FUNCTION_BLOCK AI_LAST_2 (* MERGE 2 AI in 1 AI (LAST WRITER WINS, generic FB) - welcher Socket zuletzt geschrieben hat, gewinnt und wird sofort an OUT durchgereicht *)
  (* Standard: 61499-2; Description: Copyright (c) 2026 Meisterschulen am Ostbahnhof This program and the accompanying materials are made available under the terms of the Eclipse Public License 2.0 which is available at https://www.eclipse.org/legal/epl-2.0/ SPDX-License-Identifier: EPL-2.0 *)
  (* Version 1.1, 2026-11-06, Franz Höpfinger, Meisterschulen am Ostbahnhof, generic FB GEN_AI_LAST (N Sockets), Verhalten in FORTE *)
  (* Version 1.0, 2026-08-31, Franz Höpfinger, Meisterschulen am Ostbahnhof, generic 2-way AI last-writer-wins merge, plain BasicFB (like E_D_FF/E_SR) instead of wiring F_SEL/E_RS inline every time - whichever Socket's own event fires IS the last-writer signal, no SR-latch needed *)
  PACKAGE adapter::events::unidirectional;
  IMPORT eclipse4diac::core::GenericClassName;
  {SET_ATTRIBUTE(eclipse4diac::core::GenericClassName, 'GEN_AI_LAST')}
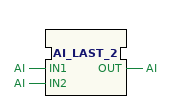
  SOCKETS
    IN1 : adapter::types::unidirectional::AI;
    IN2 : adapter::types::unidirectional::AI;
  END_SOCKETS
  PLUGS
    OUT : adapter::types::unidirectional::AI;
  END_PLUGS
END_FUNCTION_BLOCK
